TYPE ST_ModeOutputs :
STRUCT
    experimentActiveOut : BOOL;
    preArmOut : BOOL;
    resetOut : BOOL;
    enableCurrentOut : BOOL;
END_STRUCT
END_TYPE

(* stored: Version 1.1.0.1
   DUT ST_ModeOutputs: Id {0C45F671-C742-46B3-AF73-83D21687E3C8} *)
